Fanuc KAREL source: KA00185.KL

PROGRAM KA00185
%NOLOCKGROUP
VAR
  SRC: ARRAY[4] OF BYTE
  DST: ARRAY[4] OF BYTE
BEGIN
  DST = SRC
END KA00185
